ABB RobotStudio station: Pr▀ctica5_B.rspag

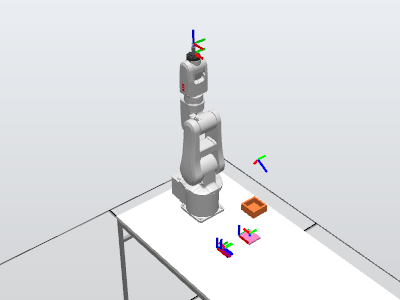
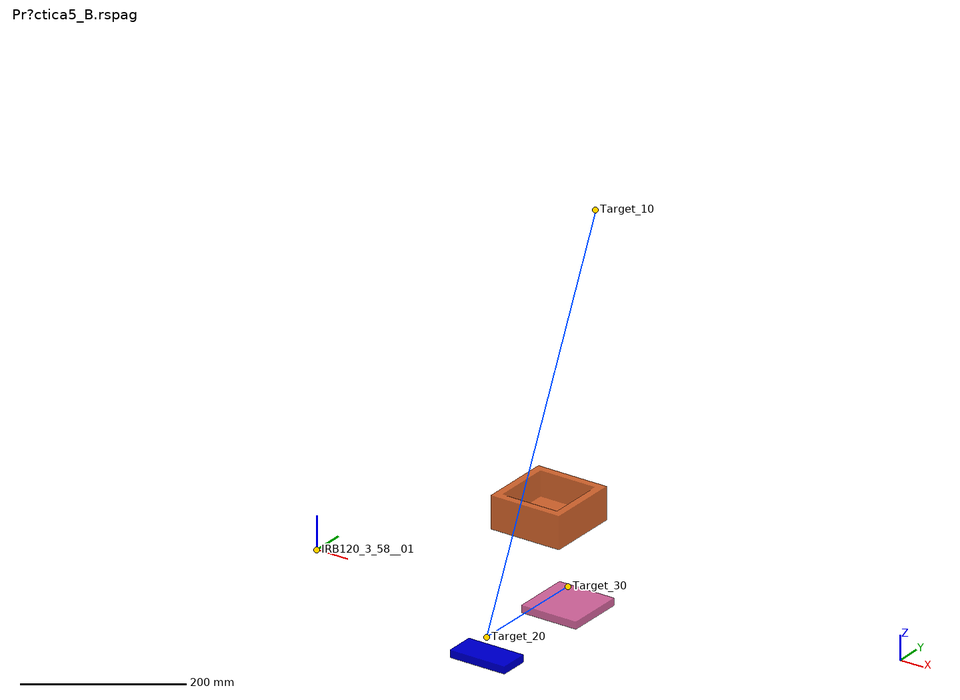
[picture v1: parts stored in the station drawn from their meshes, with robot base, taught points and paths (robot models come from the ABB library and are not in the file)]
--- station ---
Station Prßctica5_B (saved by RobotStudio 25.2.11220.0)
Controller Controlador2, task T_ROB1: task frame (RAPID world) sits at (0, 0, 670) mm in the station
Controller Controlador2
  mechanical unit ROB_1: IRB120_3_58__01, 6 joints, base frame (0, 0, 0) mm
Layout (positions relative to the parent item):
  - TVentosa [mechanism] at (-70, 0, 1604) mm
      TCP TVentosa at (0, 0, 51.19) mm
      links: Mi_herramienta
  - LogicGate [smart component, from Components\LogicGate.rslib]
      properties: Operator=NOT; Delay=0
  - LogicGate_2 [smart component, from Components\LogicGate.rslib]
      properties: Operator=AND; Delay=0
  - IRB120_3_58__01 [mechanism, from %ABB.RobotStudio.Models.IRB120%\IRB120_3_58_G_01.rslib] at (0, 0, 670) mm; joint values [0, 0, -1.5708, 0, 0, 0] (rad or m)
  - table [part, from Libraries\e293a11e-ed86-4237-866f-a9bf8f4bd145table.rslib] at (-246.62, 300, 670) mm, rotated rx 0 ry 0 rz -90 deg
  - Base2 [part], size 80 x 80 x 10 mm
  - Base1 [part], size 80 x 40 x 10 mm
  - Detacher [smart component, from Components\Detacher.rslib]
      properties: Child=Link6; KeepPosition=true
  - CollisionSensor [smart component, from Components\CollisionSensor.rslib]
      properties: Object1=TVentosa; Object2=(none); NearMiss=0.001; Part1=Mi_herramienta; Part2=Link6; CollisionType=1
    - _sensorPart_ [part]
  - Attacher_2 [smart component, from Components\Attacher.rslib]
      properties: Parent=TVentosa; Flange=0; Child=Link6; Mount=false; Offset=[0 0 0]; Orientation=[0 0 0]
  - Source_2 [smart component, from Components\Source.rslib]
      properties: Source=Pieza; Copy=(none); Parent=(none); Position=[0.34 -0.13 0.68]; Orientation=[0 0 0]; Transient=true; PhysicsBehavior=-1
  - SimulationEvents_2 [smart component, from Components\SimulationEvents.rslib]
  - Pieza [part] at (-70, 0, 1655.19) mm, size 60 x 20 x 20 mm
  - Basura [part], size 100 x 100 x 45 mm
  - LogicGate_4 [smart component, from Components\LogicGate.rslib]
      properties: Operator=AND; Delay=0
  - LogicGate_5 [smart component, from Components\LogicGate.rslib]
      properties: Operator=AND; Delay=0
  - Attacher_3 [smart component, from Components\Attacher.rslib]
      properties: Parent=TVentosa; Flange=0; Child=Link6; Mount=false; Offset=[0 0 0]; Orientation=[0 0 0]
  - CollisionSensor_2 [smart component, from Components\CollisionSensor.rslib]
      properties: Object1=TVentosa; Object2=(none); NearMiss=0.001; Part1=Mi_herramienta; Part2=Link6; CollisionType=1
    - _sensorPart_ [part]
  - LogicGate_6 [smart component, from Components\LogicGate.rslib]
      properties: Operator=AND; Delay=0
  - Detacher_2 [smart component, from Components\Detacher.rslib]
      properties: Child=Link6; KeepPosition=true
  - LogicGate_9 [smart component, from Components\LogicGate.rslib]
      properties: Operator=NOT; Delay=0
  - Sink [smart component, from Components\Sink.rslib]
      properties: Object=Link6
  - Pieza_2 [part]
  - Pieza_3 [part]
  - Pieza_4 [part]
  - Pieza_5 [part]
  - LogicGate_10 [smart component, from Components\LogicGate.rslib]
      properties: Operator=AND; Delay=0
  - LogicGate_11 [smart component, from Components\LogicGate.rslib]
      properties: Operator=NOT; Delay=0
  - LogicGate_12 [smart component, from Components\LogicGate.rslib]
      properties: Operator=NOT; Delay=0
Attachment: TVentosa is attached to IRB120_3_58__01 / Link6
Attachment: Base2 is attached to Base1
Attachment: Base1 is attached to table
Attachment: Pieza is attached to TVentosa / Mi_herramienta
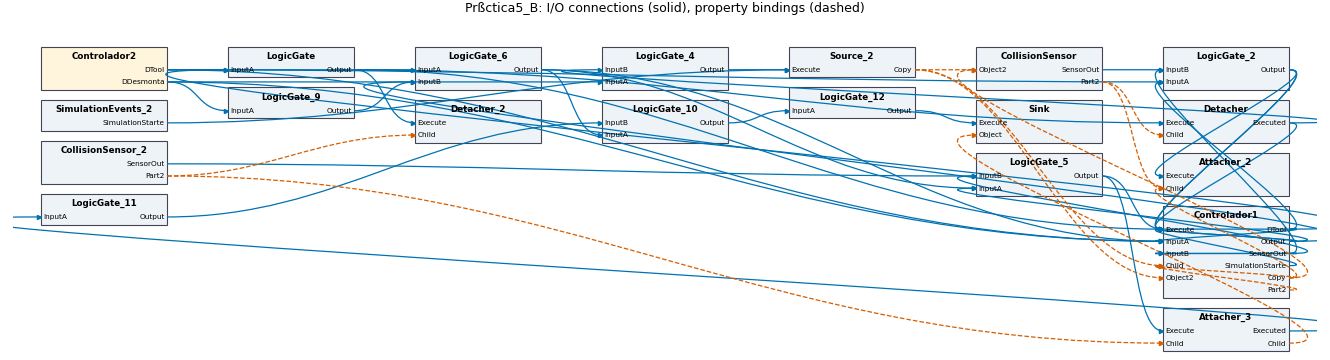
Station logic (signal -> signal, property => property):
  Controlador1.DTool -> Attacher.Execute
  Controlador1.DTool -> LogicGate_2.InputA
  LogicGate_2.Output -> Detacher.Execute
  Controlador1.DTool -> LogicGate.InputA
  LogicGate.Output -> Detacher.Execute
  CollisionSensor.SensorOut -> LogicGate_2.InputB
  Controlador1.DTool -> LogicGate_2.InputA
  LogicGate_2.Output -> Attacher.Execute
  Controlador2.DTool -> LogicGate.InputA
  LogicGate.Output -> Detacher.Execute
  Controlador2.DTool -> LogicGate_2.InputA
  LogicGate_2.Output -> Attacher.Execute
  Detacher.Executed -> Source.Execute
  SimulationEvents.SimulationStarted -> Source.Execute
  CollisionSensor.SensorOut -> LogicGate_2.InputB
  SimulationEvents_2.SimulationStarted -> Source_2.Execute
  LogicGate_2.Output -> Attacher_2.Execute
  Controlador2.DTool -> LogicGate_3.InputA
  CollisionSensor_3.SensorOut -> LogicGate_3.InputB
  LogicGate_3.Output -> Attacher_4.Execute
  CollisionSensor_4.SensorOut -> LogicGate_3.InputB
  Detacher.Executed -> LogicGate_4.InputB
  LogicGate_4.Output -> Source_2.Execute
  CollisionSensor_5.SensorOut -> LogicGate_5.InputB
  LogicGate_5.Output -> Attacher_5.Execute
  Controlador2.DDesmonta -> LogicGate_4.InputA
  CollisionSensor_2.SensorOut -> LogicGate_5.InputB
  LogicGate_5.Output -> Attacher_3.Execute
  Controlador2.DTool -> LogicGate_6.InputA
  LogicGate_6.Output -> LogicGate_7.InputA
  LogicGate_7.Output -> LogicGate_5.InputA
  LogicGate_6.Output -> LogicGate_5.InputA
  Controlador2.DDesmonta -> LogicGate_8.InputA
  LogicGate_8.Output -> LogicGate_6.InputB
  LogicGate.Output -> Detacher_2.Execute
  Controlador2.DDesmonta -> LogicGate_9.InputA
  LogicGate_9.Output -> LogicGate_6.InputB
  Attacher_3.Executed -> LogicGate_11.InputA
  LogicGate_11.Output -> LogicGate_10.InputB
  LogicGate_6.Output -> LogicGate_10.InputA
  LogicGate_10.Output -> LogicGate_12.InputA
  LogicGate_12.Output -> Sink.Execute
  Source.Copy => Attacher.Child
  Source.Copy => CollisionSensor.Object2
  Source.Copy => Attacher_2.Child
  Source_2.Copy => CollisionSensor.Object2
  Source_2.Copy => CollisionSensor_4.Object2
  Source_2.Copy => Attacher_4.Child
  CollisionSensor_5.Part2 => Attacher_5.Child
  CollisionSensor_2.Part2 => Attacher_3.Child
  CollisionSensor_2.Part2 => Detacher_2.Child
  CollisionSensor.Part2 => Attacher_2.Child
  CollisionSensor.Part2 => Detacher.Child
  Attacher_3.Child => Sink.Object

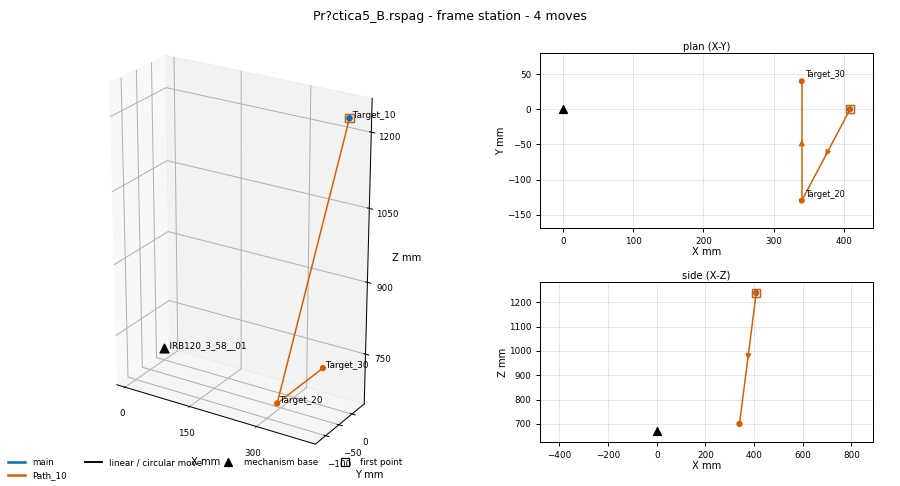
[picture p0: tool path of Pr▀ctica5_B.rspag in frame station, 4 of 16 moves have a stored position in this frame; points joined in program order, loops and branches not executed]
--- Backups/Controlador2/RAPID/TASK1/PROGMOD/CalibData.mod ---
MODULE CalibData
    PERS tooldata TVentosa:=[TRUE,[[0,0,51.19],[1,0,0,0]],[0.1,[0,0,1],[1,0,0,0],0,0,0]];
    TASK PERS wobjdata WO_Pieza:=[FALSE,TRUE,"",[[300,-150,10],[1,0,0,0]],[[20,10,0],[1,0,0,0]]];
    TASK PERS wobjdata WO_Base2:=[FALSE,TRUE,"",[[300,-150,10],[1,0,0,0]],[[0,150,0],[1,0,0,0]]];
ENDMODULE

--- Backups/Controlador2/RAPID/TASK1/PROGMOD/Module1.mod ---
MODULE Module1
    CONST robtarget Target_10:=[[408.685,0,568.405],[0.5,0,0.866025404,0],[0,0,0,0],[9E+09,9E+09,9E+09,9E+09,9E+09,9E+09]];
    CONST robtarget Target_20:=[[19.999989664,10.000006428,19.999948885],[-0.000000013,0,1,0.000000005],[-1,0,-1,0],[9E+09,9E+09,9E+09,9E+09,9E+09,9E+09]];
    CONST robtarget Target_30:=[[40,40,20],[0,0,1,0],[0,0,0,0],[9E+09,9E+09,9E+09,9E+09,9E+09,9E+09]];
    VAR num h;
    CONST jointtarget JHome:=[[0,0,-90,0,0,0],[9E+09,9E+09,9E+09,9E+09,9E+09,9E+09]];

    ! Variables Parte B
    VAR num plantas_actuales;
    VAR num plantas_nuevas;
    ! Punto de basura expresado en wobj0
    VAR robtarget Target_Basura;

    ! Medidas de la pieza (cambiar para el robot real)
    PERS num ancho_pieza:=20;
    PERS num alto_pieza:=20;

    !***********************************************************
    !
    ! Módulo:  Module1
    !
    ! Descripción: Paletizado Parte B - Torre adaptable
    !              Pick/Place genéricos (posición + workobject)
    !
    ! Autor: Javier
    !
    ! Versión: 7.0
    !
    !***********************************************************

    PROC main()
        VAR num num_pieza;
        VAR robtarget pos_pieza;

        Initialize;
        MoveJ Target_10,v200,z100,TVentosa\WObj:=wobj0;

        SetDO DDesmonta,0;

        WHILE DFin=0 DO

            TPReadNum plantas_nuevas,"Introduce el número de plantas:";

            IF plantas_nuevas>plantas_actuales THEN
                ! ---- CONSTRUCCIÓN ----
                SetDO DDesmonta,1;
                num_pieza:=plantas_actuales*4;

                WHILE DFin=0 AND num_pieza<plantas_nuevas*4 DO
                    IF DPieza=1 THEN
                        ! Coger pieza generada (en WO_Pieza)
                        Pick Target_20,WO_Pieza;
                        ! Colocar en la torre (en WO_Base2)
                        pos_pieza:=calcula_posicion(num_pieza);
                        Place pos_pieza,WO_Base2;
                        num_pieza:=num_pieza+1;
                    ENDIF
                ENDWHILE

                plantas_actuales:=plantas_nuevas;
                SetDO DDesmonta,0;

            ELSEIF plantas_nuevas<plantas_actuales THEN
                ! ---- DESMONTAJE ----
                SetDO DDesmonta,0;
                num_pieza:=plantas_actuales*4-1;

                WHILE num_pieza>=plantas_nuevas*4 DO
                    ! Coger pieza de la torre (en WO_Base2)
                    pos_pieza:=calcula_posicion(num_pieza);
                    Pick pos_pieza,WO_Base2;
                    ! Dejar en la basura (en WO_Base2)
                    Place Target_Basura,WO_Base2;
                    num_pieza:=num_pieza-1;
                ENDWHILE

                plantas_actuales:=plantas_nuevas;

            ENDIF

        ENDWHILE

        MoveAbsJ JHome,v150,z200,TVentosa\WObj:=wobj0;
    ENDPROC

    FUNC robtarget calcula_posicion(num num_pieza)
        VAR robtarget punto;
        VAR num tipo;
        VAR num piso;
        VAR num z_planta;

        tipo:=num_pieza MOD 4;
        piso:=num_pieza DIV 4;
        z_planta:=piso*2*alto_pieza;

        TEST tipo
        CASE 0:
            punto:=Offs(Target_30,0,ancho_pieza,z_planta);
        CASE 1:
            punto:=Offs(Target_30,0,-ancho_pieza,z_planta);
        CASE 2:
            punto:=Offs(Target_30,ancho_pieza,0,z_planta+alto_pieza);
            punto.rot:=OrientZYX(90,0,180);
        CASE 3:
            punto:=Offs(Target_30,-ancho_pieza,0,z_planta+alto_pieza);
            punto.rot:=OrientZYX(90,0,180);
        DEFAULT:
            punto:=Target_30;
        ENDTEST

        RETURN punto;
    ENDFUNC

    PROC Initialize()
        h:=0;
        plantas_actuales:=0;
        plantas_nuevas:=0;
        SetDO DTool,0;
        ! Punto de basura relativo a WO_Base2
        Target_Basura.trans.x:=-100;
        Target_Basura.trans.y:=200;
        Target_Basura.trans.z:=20;
        Target_Basura.rot:=[0,0,1,0];
        Target_Basura.robconf:=[0,0,0,0];
        Target_Basura.extax:=[9E+09,9E+09,9E+09,9E+09,9E+09,9E+09];
    ENDPROC

    PROC Pick(robtarget posicion,PERS wobjdata wobj_uso)
        ConfJ\Off;
        ConfL\Off;
        ! Aproximación 100mm arriba
        MoveJ Offs(posicion,0,0,100),v500,z50,TVentosa\WObj:=wobj_uso;
        ! Aproximación 50mm arriba
        MoveJ Offs(posicion,0,0,50),v200,z10,TVentosa\WObj:=wobj_uso;
        ! Punto destino
        MoveJ posicion,v100,fine,TVentosa\WObj:=wobj_uso;
        ! Coger
        SetDO DTool,1;
        WaitTime 0.3;
        ! Subir
        MoveJ Offs(posicion,0,0,50),v200,z10,TVentosa\WObj:=wobj_uso;
        MoveJ Offs(posicion,0,0,100),v500,z50,TVentosa\WObj:=wobj_uso;
        ConfJ\On;
        ConfL\On;
    ENDPROC

    PROC Place(robtarget posicion,PERS wobjdata wobj_uso)
        ConfJ\Off;
        ConfL\Off;
        ! Aproximación 100mm arriba
        MoveJ Offs(posicion,0,0,100),v500,z50,TVentosa\WObj:=wobj_uso;
        ! Aproximación 50mm arriba
        MoveJ Offs(posicion,0,0,50),v200,z10,TVentosa\WObj:=wobj_uso;
        ! Punto destino
        MoveJ posicion,v100,fine,TVentosa\WObj:=wobj_uso;
        ! Soltar
        SetDO DTool,0;
        WaitTime 0.3;
        ! Subir
        MoveJ Offs(posicion,0,0,50),v200,z10,TVentosa\WObj:=wobj_uso;
        MoveJ Offs(posicion,0,0,100),v500,z50,TVentosa\WObj:=wobj_uso;
        ConfJ\On;
        ConfL\On;
    ENDPROC

    PROC Path_10()
        MoveJ Target_10,v200,z100,TVentosa\WObj:=wobj0;
        MoveL Target_20,v200,fine,TVentosa\WObj:=WO_Pieza;
        MoveL Target_30,v200,z100,TVentosa\WObj:=WO_Base2;
        MoveAbsJ JHome,v200,z100,TVentosa\WObj:=WO_Pieza;
    ENDPROC

ENDMODULE

--- Backups/Controlador2/SYSPAR/EIO.cfg ---
EIO:CFG_1.0:6:1::
#
EIO_SIGNAL:

      -Name "DFin" -SignalType "DI"

      -Name "DTool" -SignalType "DO"

      -Name "DPieza" -SignalType "DI"

      -Name "DDesmonta" -SignalType "DO"
